// TIA Portal V20 export
// export: Created 2026-10-12T05:00:28.5696988Z, ExportSetting WithDefaults, DisplayName Totally Integrated Automation Portal, DisplayVersion V20, DisplayName TIA Portal Openness, DisplayVersion V20, DisplayName TIA Portal Teamcenter Gateway, DisplayVersion V20, DisplayName TIA Portal Version Control Interface, DisplayVersion V20, DisplayName SINAMICS Startdrive Advanced, DisplayVersion V20 SP1 Update 2, DisplayName SINAMICS Startdrive G110M, G120, G120C, G120D, G120P, G115D, DisplayVersion V20 SP1 Update 2, DisplayName SINAMICS Startdrive G130, G150, S120, S150, SINAMICS MV, G220, S200, S210, DisplayVersion V20 SP1 Update 2, DisplayName STEP 7 Professional, DisplayVersion V20, DisplayName STEP 7 Safety, DisplayVersion V20, DisplayName WinCC Basic/Comfort/Advanced, DisplayVersion V20, DisplayName WinCC Professional, DisplayVersion V20, DisplayName WinCC Unified, DisplayVersion V20
FUNCTION "FRK_AccessPolicySave" : Void   // FC59, SCL
{ S7_Optimized_Access := 'TRUE' }
VERSION : 0.1
// stored: AutoNumber true, IsIECCheckEnabled false, SetENOAutomatically false, UDAEnableTagReadback false
   VAR_INPUT
      Scope : String;
   END_VAR
   VAR_IN_OUT
      Access : "FRK_Access";
   END_VAR
BEGIN

   IF #Access.PolicySlot < 1 OR #Access.PolicySlot > 2 THEN
       RETURN;
   END_IF;
   IF #Scope = '' OR NOT "FRK_AccessPolicyShape"(Policy := #Access.Policy) THEN
       #Access.PolicyLost := TRUE;
       RETURN;
   END_IF;
   "FRK_AccessPolicies".Rows[#Access.PolicySlot].SchemaVersion := 1;
   "FRK_AccessPolicies".Rows[#Access.PolicySlot].Scope := #Scope;
   "FRK_AccessPolicies".Rows[#Access.PolicySlot].Generation := "FRK_AccessNext"(Previous := "FRK_AccessPolicies".Rows[#Access.PolicySlot].Generation);
   "FRK_AccessPolicies".Rows[#Access.PolicySlot].Policy := #Access.Policy;
   "FRK_AccessPolicies".Rows[#Access.PolicySlot].Checksum := "FRK_AccessPolicyCrc"(Image := "FRK_AccessPolicies".Rows[#Access.PolicySlot]);
END_FUNCTION
